(* IEC 61131-3 sources: llm-plc-st-eval/data/definitivo/claude-sonnet-4-6/C8/few_shot, 3 files *)

(* ---- ejec_1.st ---- *)
```pascal
FUNCTION_BLOCK FB_Valvula
VAR_INPUT
    nivelAlto : BOOL; (* Contacto NA: activa el temporizador *)
END_VAR
VAR_OUTPUT
    valvula : BOOL; (* Bobina: activada tras retardo *)
END_VAR
VAR
    T1 : TON; (* Temporizador a la conexión, PT = 5 s *)
END_VAR

(* Rama 1: nivelAlto alimenta la entrada IN del TON T1 *)
T1(IN := nivelAlto, PT := T#5S);

(* Rama 2: la salida Q de T1 alimenta la bobina valvula *)
valvula := T1.Q;

END_FUNCTION_BLOCK
```

(* ---- ejec_2.st ---- *)
```st
FUNCTION_BLOCK FB_Valvula
VAR_INPUT
    nivelAlto : BOOL; (* Contacto NA que activa el temporizador *)
END_VAR
VAR_OUTPUT
    valvula : BOOL; (* Bobina activada tras el retardo *)
END_VAR
VAR
    T1 : TON; (* Temporizador a la conexión, retardo de 5 s *)
END_VAR

(* Rama 1: nivelAlto alimenta la entrada IN del TON T1 *)
T1(IN := nivelAlto, PT := T#5S);

(* Rama 2: T1.Q (contacto NA) alimenta la bobina valvula *)
valvula := T1.Q;

END_FUNCTION_BLOCK
```

(* ---- ejec_3.st ---- *)
```st
FUNCTION_BLOCK FB_Valvula
VAR_INPUT
    nivelAlto : BOOL; (* Contacto NA: activa el temporizador *)
END_VAR
VAR_OUTPUT
    valvula : BOOL; (* Bobina: se activa cuando T1.Q es TRUE *)
END_VAR
VAR
    T1 : TON; (* Temporizador a la conexión, tiempo preestablecido 5 s *)
END_VAR

(* Rama 1: nivelAlto alimenta la entrada IN del TON T1 *)
T1(IN := nivelAlto, PT := T#5S);

(* Rama 2: la salida Q de T1 alimenta la bobina valvula *)
valvula := T1.Q;
END_FUNCTION_BLOCK
```
